{attribute 'qualified_only'}
{attribute 'strict'}
TYPE E_EventSeverity :
(
    Error,
    Warning,
    Info
);
END_TYPE

(* stored: Version 1.1.0.1, ProductVersion 3.1.4026.18
   DUT E_EventSeverity: Id {108656a3-bb94-49ab-be2d-18f5161d1fdc} *)
